// TIA Portal V21 export
// export: Created 2026-11-10T22:46:46.7831663Z, ExportSetting WithDefaults, DisplayName Totally Integrated Automation Portal, DisplayVersion V21 Update 3, DisplayName STEP 7 Professional, DisplayVersion V21 Update 3, DisplayName STEP 7 Safety, DisplayVersion V21, DisplayName Tech WebApplication, DisplayVersion V21, DisplayName WinCC Basic/Comfort/Advanced, DisplayVersion V21 Update 3, DisplayName WinCC Unified, DisplayVersion V21 Update 3
FUNCTION "FC_Ton" : Void   // FC1, SCL
{ S7_Optimized_Access := 'TRUE' }
VERSION : 0.1
// stored: AutoNumber true, IsIECCheckEnabled false, SetENOAutomatically false, UDAEnableTagReadback false
   VAR_INPUT
      start : Bool;
   END_VAR
   VAR_OUTPUT
      q : Bool;
   END_VAR
BEGIN
   "DBTon".TON(IN := #start, PT := T#2S);
           #q := "DBTon".Q;
END_FUNCTION
